// TwinCAT 3 PLC project slavePLC
// ProgramVersion: 3.1.4026.20
// libraries:
//   Tc2_Standard, * (Beckhoff Automation GmbH)
//   Tc2_System, * (Beckhoff Automation GmbH)
//   Tc3_Module, * (Beckhoff Automation GmbH)
//   VisuSymbols,3.5.10.0,System
// project tree:
//   / GlobalTextList.TcGTLO, PlcTask.TcTTO, Visualization Manager.TcVMO (not stored)
//   GVLs/ GVLSlave.TcGVL, ImagePoolCar.TcIPO (not stored)
//   POUs/ CarContorl.TcPOU, LampDelay.TcPOU, LampSlave.TcPOU, LongHandshake.TcPOU, MAIN.TcPOU, RunSlave.TcPOU, ShortHandshake.TcPOU, SlaveHandeshake.TcPOU
//   VISUs/ VisualizationSlave.TcVIS
// (motion and I/O tree: see PLC project studentplc)
// real-time tasks:
//   TASK PlcTask: cycle T#10ms, priority 20, ADS port 350
//   TASK PlcTask1: cycle T#10ms, priority 21, ADS port 351
// variable links:
//   StudentPLC/StudentPLC Instance <-> slavePLC/slavePLC Instance
//     PlcTask Inputs/GVLStudent.ixStrobOne <-> PlcTask Outputs/GVLSlave.oxStrobOne
//     PlcTask Inputs/GVLStudent.ixStrobTwo <-> PlcTask Outputs/GVLSlave.oxStrobTwo
//     PlcTask Outputs/GVLStudent.IXButtonLong <-> PlcTask Inputs/GVLSlave.ixLong
//     PlcTask Outputs/GVLStudent.IXButtonShort <-> PlcTask Inputs/GVLSlave.ixShort
//     PlcTask Outputs/GVLStudent.oxStrobOne <-> PlcTask Inputs/GVLSlave.ixStrobOne
//     PlcTask Outputs/GVLStudent.oxStrobTwo <-> PlcTask Inputs/GVLSlave.ixStrobTwo

CONFIGURATION slavePLC
    RESOURCE PLC ON TwinCAT3
        TASK PlcTask(INTERVAL := T#10ms, PRIORITY := 21);
        PROGRAM MAIN WITH PlcTask : MAIN;
    END_RESOURCE
END_CONFIGURATION

// ---- GVLs/GVLSlave.TcGVL
{attribute 'qualified_only'}
VAR_GLOBAL
	
	// Lamp varibol
	OXLampOXOne :BOOL;
	OXLampIXOneGreen :BOOL;
	OXLampOXTwo :BOOL;
	OXLampIXTwoGreen :BOOL;
	
	//strob out
	oxStrobOne AT %Q* : BOOL ;
	oxStrobTwo AT %Q* : BOOL ;
 	//strob in
	ixStrobOne AT %I* : BOOL ;
	ixStrobTwo AT %I* : BOOL ;
	
	// Long or Short
	ixLong AT %I* : BOOL;
	ixShort AT%I* :BOOL;
	
	// car move
	OIntRedCar: INT;
	OintCopCar: INT;
END_VAR

// ---- POUs/MAIN.TcPOU
PROGRAM MAIN
VAR
END_VAR

RunSlave();

END_PROGRAM

// ---- POUs/RunSlave.TcPOU
PROGRAM RunSlave
VAR
	LampSlave_0: LampSlave;
	SlaveHandeshake_0: SlaveHandeshake;
	ixStrobOne :BOOL;
	ixStrobTwo :BOOL;
	startCar: BOOL;
	carEnd: BOOL;
	CarContorl_0: CarContorl;
END_VAR

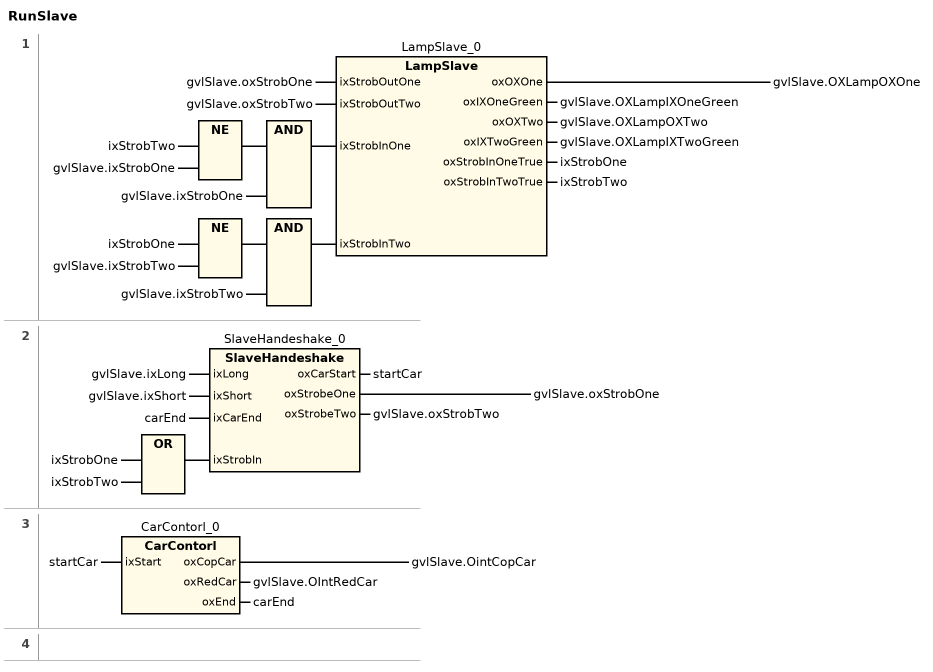
// NETWORK 1
LampSlave_0(
    ixStrobOutOne := gvlSlave.oxStrobOne,
    ixStrobOutTwo := gvlSlave.oxStrobTwo,
    ixStrobInOne := ixStrobTwo <> gvlSlave.ixStrobOne AND gvlSlave.ixStrobOne,
    ixStrobInTwo := ixStrobOne <> gvlSlave.ixStrobTwo AND gvlSlave.ixStrobTwo,
    oxIXOneGreen => gvlSlave.OXLampIXOneGreen,
    oxOXTwo => gvlSlave.OXLampOXTwo,
    oxIXTwoGreen => gvlSlave.OXLampIXTwoGreen,
    oxStrobInOneTrue => ixStrobOne,
    oxStrobInTwoTrue => ixStrobTwo); // LampSlave
gvlSlave.OXLampOXOne := LampSlave_0.oxOXOne;

// NETWORK 2
SlaveHandeshake_0(
    ixLong := gvlSlave.ixLong,
    ixShort := gvlSlave.ixShort,
    ixCarEnd := carEnd,
    ixStrobIn := ixStrobOne OR ixStrobTwo,
    oxCarStart => startCar,
    oxStrobeTwo => gvlSlave.oxStrobTwo); // SlaveHandeshake
gvlSlave.oxStrobOne := SlaveHandeshake_0.oxStrobeOne;

// NETWORK 3
CarContorl_0(ixStart := startCar, oxRedCar => gvlSlave.OIntRedCar, oxEnd => carEnd); // CarContorl
gvlSlave.OintCopCar := CarContorl_0.oxCopCar;

// NETWORK 4

END_PROGRAM

// ---- POUs/LampSlave.TcPOU
FUNCTION_BLOCK LampSlave
VAR_INPUT
	ixStrobOutOne :BOOL; // Direct control for group One main lamp (OX1)
	ixStrobOutTwo :BOOL; // Direct control for group Two main lamp (OX2)
	
	ixStrobInOne: BOOL; // Start signal for LampDelay sequence (group One)
	ixStrobInTwo: BOOL; // Start signal for LampDelay sequence (group Two)

END_VAR
VAR_OUTPUT
	  // Group One: main lamp + 3 indicator lamps (R, B, G)
	oxOXOne :BOOL; // Main lamp (direct)
	
	oxIXOneGreen :BOOL; // Indicator Green (from LampDelay)
	
	oxOXTwo :BOOL; // Main lamp (direct)
	
	oxIXTwoGreen :BOOL; // Indicator Green (from LampDelay)
	
	oxStrobInOneTrue: BOOL; // TRUE when all three indicators (group One) are ON
	oxStrobInTwoTrue: BOOL;// TRUE when all three indicators (group Two) are ON
	
END_VAR
	
VAR
	
	LampIXOne : LampDelay; // Instance for group One sequence
	LampIXTwo : LampDelay; // Instance for group Two sequence
	
END_VAR

// ------------------------------
// Direct main-lamp control
// ------------------------------

IF ixStrobOutOne THEN
	oxOXOne := TRUE;
ELSE
	oxOXOne := FALSE;
END_IF

IF ixStrobOutTwo THEN
	oxOXTwo := TRUE;
ELSE
	oxOXTwo := FALSE;
END_IF



// ------------------------------
// Group One: delayed indicator sequence
// ------------------------------
LampIXOne(ixStart := ixStrobInOne);

// Map LampDelay outputs to group One indicators
oxIXOneGreen     := LampIXOne.oxLampThree; // Green
oxStrobInOneTrue := LampIXOne.oxAllLightsOn; // All indicators ON


// ------------------------------
// Group Two: delayed indicator sequence
// ------------------------------
LampIXTwo(ixStart := ixStrobInTwo);

// Map LampDelay outputs to group Two indicators
oxIXTwoGreen     := LampIXTwo.oxLampThree; // Green
oxStrobInTwoTrue := LampIXTwo.oxAllLightsOn; // All indicators ON

END_FUNCTION_BLOCK

// ---- POUs/LampDelay.TcPOU
FUNCTION_BLOCK LampDelay
VAR_INPUT
    ixStart : BOOL;      // Start command: TRUE = run "power-up" sequence; FALSE = run "power-down" sequence
END_VAR
VAR_OUTPUT
    oxLampThree    : BOOL; // Output: Lamp 3 on/off
    oxAllLightsOn  : BOOL; // TRUE when all three lamps are on
END_VAR
VAR
    t      : TON;             // TON timer instance (non-retentive on IN falling edge)
    step   : INT := 0;        // State machine step
    delay  : TIME := T#2S;    // Delay duration used between steps
    tStart : BOOL;            // Timer IN signal (acts like a "strobe" to start the TON)
    tEnd   : BOOL;            // TRUE when timer has elapsed (t.Q)
END_VAR


//_______________________________________________________________________________________________
// LampDelay is a step-sequenced (state machine) controller that turns on three lamps
// one BY one with a fixed delay between each stage when ixStart is TRUE. 
// When ixStart goes FALSE, it turns the lamps off again in reverse order, also with delays. 
// A TON timer (t) provides the per-step delay. oxAllLightsOn is TRUE once all three lamps are on.
//_______________________________________________________________________________________________


// ------------------------------
// State machine for sequenced on/off with delays
// ------------------------------
CASE step OF

    0: // Idle/reset: all lamps off, wait for start
        oxLampThree    := FALSE;
        oxAllLightsOn  := FALSE;
        IF ixStart THEN
            // Start power-up sequence: immediately turn on Lamp 1 and start delay
            tStart    := TRUE;                  // Start the TON for the next step delay
			t(IN := tStart, PT := delay);
            step      := 20;
        END_IF


    20: // After Lamp 2 is on, wait delay, then turn on Lamp 3
        IF tEnd THEN
            tStart := FALSE;                   // Reset TON input before next start
            t(IN := tStart, PT := delay);
            oxLampThree := TRUE;
            step := 30;
        END_IF

    30: // All three lamps are on; assert "all on" and wait for stop command
        oxAllLightsOn := TRUE;
        IF NOT ixStart THEN
            // Begin power-down sequence after stop command
            tStart := TRUE;                    // Start delay before turning lamps off
            t(IN := tStart, PT := delay);
            step := 60;
        END_IF


    60: // Wait delay, then turn off Lamp 1 and return to idle
        IF tEnd THEN
            oxLampThree := FALSE;
			tStart := FALSE;
			t(IN := tStart,  PT := delay);
            step := 0;                         // Back to idle
        END_IF

END_CASE

// ------------------------------
// Timer execution (must be called each cycle)
// ------------------------------
t(IN := tStart, PT := delay);  // Evaluate TON with current IN/PT
tEnd := t.Q;                   // Timer done flag for step logic

END_FUNCTION_BLOCK

// ---- POUs/SlaveHandeshake.TcPOU
FUNCTION_BLOCK SlaveHandeshake
VAR_INPUT
	ixLong :BOOL;
	ixShort :BOOL;
	ixCarEnd: BOOL;
	ixStrobIn :BOOL; 
END_VAR
VAR_OUTPUT
	oxCarStart: BOOL;
	oxStrobeOne : BOOL;
    oxStrobeTwo : BOOL;
END_VAR
VAR
	
	long : LongHandshake;
	short : ShortHandshake;  
	oxStrobeOneShort : BOOL;
	oxStrobeOneLong : BOOL;
	oxCarStartLong: BOOL;
	oxCarStartShort: BOOL;
	step : INT := 0;
	waitLong : BOOL;
	waitShort: BOOL;
END_VAR

// ------------------------------
// State selector: choose which handshake to run
// ------------------------------
CASE step OF

    0: // IDLE: wait for a mode selection
        // NOTE: If both ixLong and ixShort are TRUE, long wins here.
        IF ixLong THEN
            step := 10;
        ELSIF ixShort THEN
            step := 20;
        END_IF

    10: // RUN LONG HANDSHAKE
        long(ixStart := ixCarEnd, ixStrobIn := ixStrobIn);

        // Map long handshake outputs to locals
        oxStrobeOneLong := long.oxStrobeOne;
        oxStrobeTwo     := long.oxStrobeTwo;  // direct passthrough (long only)
        oxCarStartLong  := long.oxStart;
        waitLong        := long.oxwait;

        // When long handshake reports idle, return to IDLE
        IF waitLong THEN
            step := 0;
        END_IF

    20: // RUN SHORT HANDSHAKE
        short(ixStart := ixCarEnd, ixStrobIn := ixStrobIn);

        // Map short handshake outputs to locals
        oxStrobeOneShort := short.oxStrobe;
        oxCarStartShort  := short.oxStart;
        waitShort        := short.oxwait;     // FIX: lowercase 'short'

        // When short handshake reports idle, return to IDLE
        IF waitShort THEN
            step := 0;
        END_IF

END_CASE


// ------------------------------
// Common output mapping
// ------------------------------

// Car start/ack goes TRUE if either handshake asserts it
IF oxCarStartShort OR oxCarStartLong THEN 
	oxCarStart := TRUE; 
ELSE 
	oxCarStart := FALSE; 
END_IF

// Primary strobe is TRUE if either handshake asserts it
IF oxStrobeOneShort OR oxStrobeOneLong THEN
	oxStrobeOne := TRUE; 
ELSE 
	oxStrobeOne := FALSE; 
END_IF

END_FUNCTION_BLOCK

// ---- POUs/LongHandshake.TcPOU
FUNCTION_BLOCK LongHandshake
VAR_INPUT
    ixStart   : BOOL; // From Master: start command ("execute now")
    ixStrobIn : BOOL; // From Master: strobe/ack line used through the long handshake
END_VAR
VAR_OUTPUT
    oxStart     : BOOL; // To Master: Slave "start request" (go-high to request start)
    oxStrobeOne : BOOL; // To Master: first Slave strobe (ack for initial Master strobe)
    oxStrobeTwo : BOOL; // To Master: second Slave strobe (ack after start)
    oxwait      : BOOL; // TRUE when idle/waiting; FALSE during handshake
END_VAR
VAR
    step : INT := 0;     // State machine step
END_VAR

CASE step OF

    0:  // IDLE: reset strobes, signal wait, and watch for Master strobe
        oxStrobeOne := FALSE;
        oxStrobeTwo := FALSE;
        oxStart     := FALSE;   // Ensure start request is low in idle
        oxwait      := TRUE;

        IF ixStrobIn THEN
            // Master raised strobe → acknowledge with Slave strobe one
            oxStrobeOne := TRUE;
            oxwait      := FALSE;
            step        := 10;
        END_IF

    10: // HOLD STROBE ONE until Master drops its strobe
        oxStrobeOne := TRUE;

        IF NOT ixStrobIn THEN
            // Master dropped strobe → drop Slave strobe one and move on
            oxStrobeOne := FALSE;
            step        := 20;
        END_IF

    20: // REQUEST START: raise oxStart to ask Master to start
        oxStart := TRUE;        // Keep high until Master issues ixStart

        IF ixStart THEN
            // Start received → drop request and raise second strobe
            oxStart     := FALSE;
            oxStrobeTwo := TRUE;
            step        := 30;
        END_IF

    30: // HOLD STROBE TWO until Master acknowledges (raises its strobe)
        oxStrobeTwo := TRUE;

        IF ixStrobIn THEN
            // Master acknowledged → drop strobe two and wait for final low
            oxStrobeTwo := FALSE;
            step        := 40;
        END_IF

    40: // WAIT FOR MASTER TO RETURN LOW to complete the cycle
        oxStrobeTwo := FALSE;

        IF NOT ixStrobIn THEN
            // Handshake finished → back to idle
            step := 0;
        END_IF

END_CASE

END_FUNCTION_BLOCK

// ---- POUs/ShortHandshake.TcPOU
FUNCTION_BLOCK ShortHandshake
VAR_INPUT
    ixStart   : BOOL; // Input from Master: start command ("execute now")
    ixStrobIn : BOOL; // Input from Master: strobe/trigger to initiate the handshake
END_VAR

VAR_OUTPUT
    oxStart  : BOOL; // Output to Master: "acknowledge/ready" from Slave
    oxStrobe : BOOL; // Output to Master: Slave strobe/confirmation during handshake
    oxwait   : BOOL; // Output: TRUE when Slave is idle/waiting
END_VAR

VAR
    step : INT := 0; // State machine step
END_VAR


// ------------------------------
// Short handshake sequence (Slave side)
// Step 0: Idle, waiting for Master strobe (ixStrobIn = TRUE)
// Step 10: Acknowledge/ready (oxStart = TRUE) until Master issues start (ixStart = TRUE)
// Step 20: Slave strobe (oxStrobe = TRUE) until Master drops its strobe (ixStrobIn = FALSE)
// ------------------------------
CASE step OF

    0:  // IDLE: reset all signals, wait for Master strobe
        oxStrobe := FALSE;
        oxStart  := FALSE;
        oxwait   := TRUE;

        IF ixStrobIn THEN
            // Master raised strobe → acknowledge and go to READY
            oxStart := TRUE;
            oxwait  := FALSE;
            step    := 10;
        END_IF

    10: // READY: wait for Master start command
        oxStart := TRUE;   // Keep acknowledge high

        IF ixStart THEN
            // Master gave start → drop ack and raise Slave strobe
            oxStart  := FALSE;
            oxStrobe := TRUE;
            step     := 20;
        END_IF

    20: // SLAVE STROBE: hold until Master drops its strobe
        oxStrobe := TRUE;

        IF NOT ixStrobIn THEN
            // Master strobe dropped → finish cycle and return to idle
            oxStrobe := FALSE;
            step     := 0;
        END_IF

END_CASE

END_FUNCTION_BLOCK

// ---- POUs/CarContorl.TcPOU
FUNCTION_BLOCK CarContorl
VAR_INPUT
    ixStart : BOOL;         // Start signal: TRUE = run sequence, FALSE = reset
END_VAR
VAR_OUTPUT
    oxCopCar : INT;         // Position counter for Cop car (moves negative)
    oxRedCar : INT;         // Position counter for Red car (moves negative)
    oxEnd    : BOOL;        // TRUE when both cars reach their thresholds
END_VAR
VAR
    step   : INT := 0;      // Step in the state machine
    t      : TON;           // TON timer instance (1s delay)
    delay  : TIME := T#1S;  // Delay interval
    tStart : BOOL;          // TON input (used as strobe to retrigger timer)
    tEnd   : BOOL;          // TON output (TRUE when delay time has passed)
END_VAR

//_______________________________________________________________________________________________________________
// CarContorl is a simple state machine that simulates two “cars” moving when the start signal (ixStart) is TRUE.
// Every second, the Cop car counter decreases by 2 and the Red car counter decreases by 3.
// When both cars pass their thresholds (Cop ≤ −800 and Red ≤ −1000), the output oxEnd is set TRUE.
// If ixStart goes FALSE, everything resets to the initial state.
//______________________________________________________________________________________________________________

CASE step OF

    0:  // IDLE/RESET: clear outputs and wait for start
        oxEnd    := FALSE;
        oxCopCar := 0;
        oxRedCar := 0;

        IF ixStart THEN
            tStart := TRUE;                // Start the first delay
            t(IN := tStart, PT := delay);
            step := 1;
        END_IF

    1:  // UPDATE POSITION: decrement both cars each cycle
        oxCopCar := oxCopCar - 2;          // Cop car moves -2 per step
        oxRedCar := oxRedCar - 3;          // Red car moves -3 per step

        IF tEnd THEN                       // After 1 second → go to check
            step := 10;
        END_IF

    10: // CHECK GOALS: have both thresholds been reached?
        IF (oxCopCar <= -800) AND (oxRedCar <= -1000) THEN
            oxEnd := TRUE;                 // Both goals reached → finish
            step  := 20;
        ELSE
            // Not yet → retrigger TON for next cycle
            tStart := FALSE;               // Reset TON input
            t(IN := tStart, PT := delay);
            tStart := TRUE;                // Rising edge to retrigger TON
            t(IN := tStart, PT := delay);
            step := 1;                     // Continue updating
        END_IF

    20: // FINISHED: hold end signal until start goes low
        oxEnd := TRUE;

        IF NOT ixStart THEN                // Stop command → reset
            oxEnd := FALSE;
            step  := 0;
        END_IF

END_CASE

// ------------------------------
// Timer evaluation – must be called every cycle
// ------------------------------
t(IN := tStart, PT := delay);
tEnd := t.Q;

END_FUNCTION_BLOCK

// ---- GlobalTextList.TcGTLO
TEXTLIST GlobalTextList
  76 = "first strobe '\\n' downloaded"
  36 = 'first strobe downloaded'
  378 = 'IXOne'
  620 = 'IXTwo'
  958 = 'loading'
  923 = 'Looding'
  389 = 'Loodining'
  816 = 'OXOne'
  99 = 'OXTwo'
  160 = 'Slav PLC'
  965 = 'Slav Strob One '
  171 = 'Slav strob one send'
  590 = 'Slav strob Two send'
  605 = 'Slav strob two send'
  659 = 'Strob sent'
  46 = 'strobe downloaded'
  781 = 'Strobe downloaded'
  391 = 'strobe received'
  968 = 'Strobe received'
END_TEXTLIST

// ---- VISUs/VisualizationSlave.TcVIS
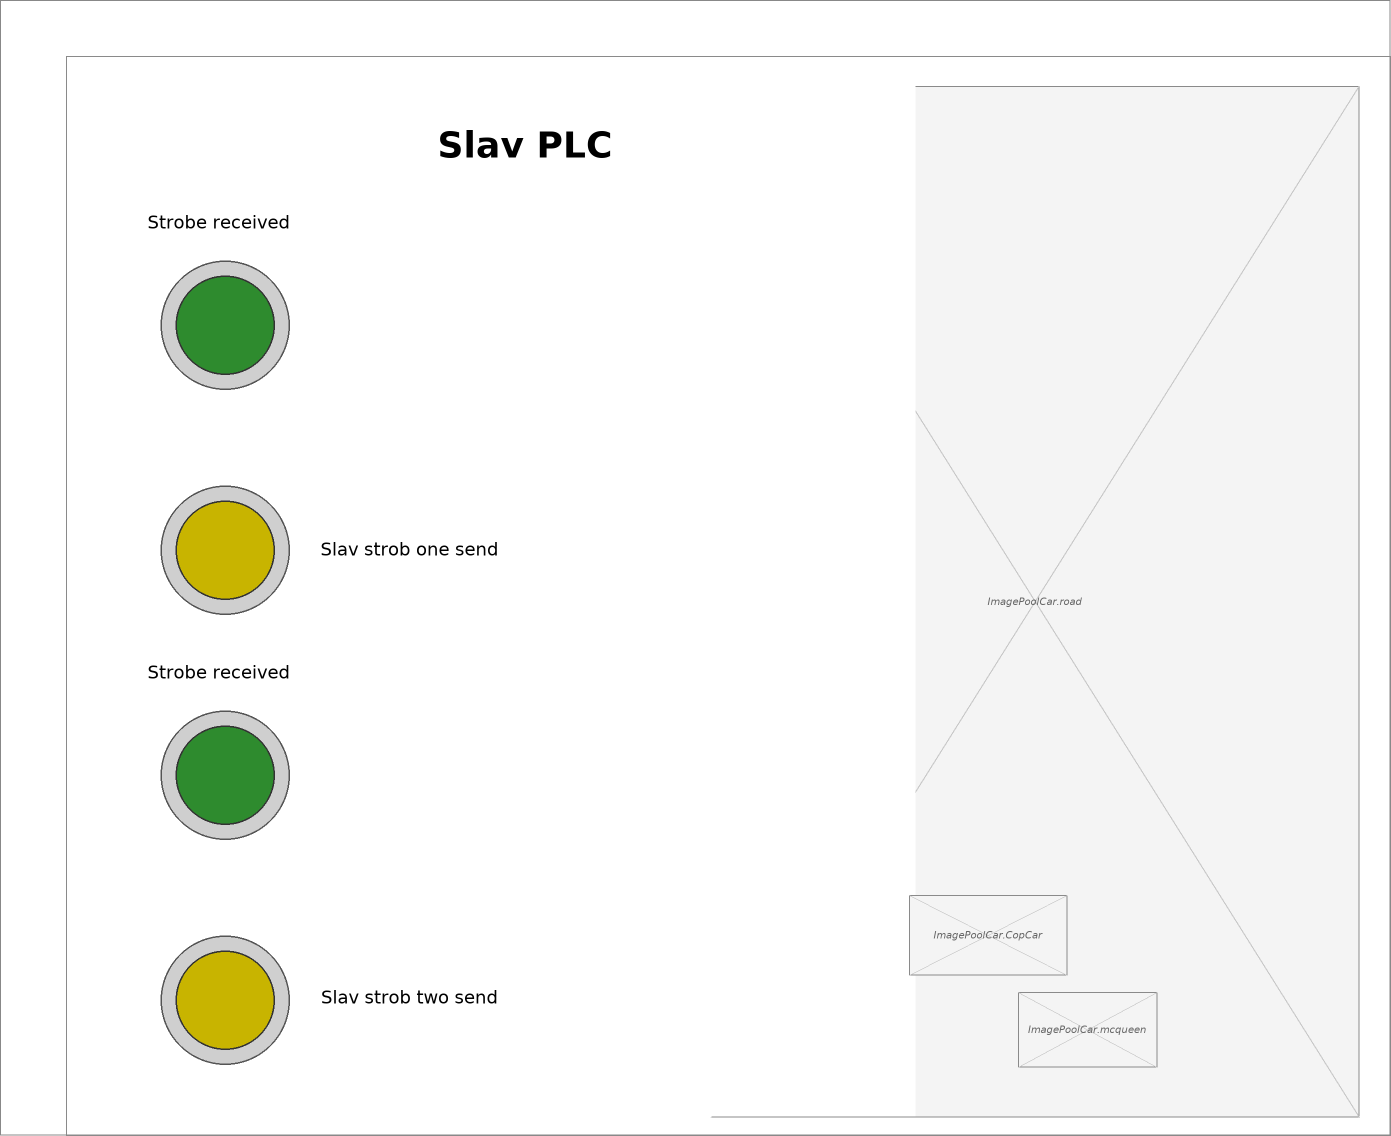
VISUALIZATION VisualizationSlave  // 1391x1136
    Frame (66,56 1325x1080)
    Image (711,86 648x1031), image: ImagePoolCar.road
    Rectangle (637,86 278x1030)
    Label (400,120 250x50), "Slav PLC"
    Lamp1 (150,250 150x150), variable: GVLSlave.OXLampIXOneGreen, style: Lamp-Lamp1-Green
    Label (100,200 238x45), "Strobe received"
    Label (300,527 219x45), "Slav strob one send"
    Lamp1 (150,475 150x150), variable: GVLSlave.OXLampOXOne, style: Lamp-Lamp1-Yellow
    Lamp1 (150,700 150x150), variable: GVLSlave.OXLampIXTwoGreen, style: Lamp-Lamp1-Green
    Lamp1 (150,925 150x150), variable: GVLSlave.OXLampOXTwo, style: Lamp-Lamp1-Yellow
    Image (1018,992 139x75), angle 90, image: ImagePoolCar.mcqueen
        p3528305787: GVLSlave.OIntRedCar
        p874137650: GVLSlave.OIntRedCar
    Image (909,895 158x80), angle 90, image: ImagePoolCar.CopCar
        p3528305787: GVLSlave.OintCopCar
        p874137650: GVLSlave.OintCopCar
    Label (300,975 219x45), "Slav strob two send"
    Label (100,650 238x45), "Strobe received"
    Label (450,650 150x30)
END_VISUALIZATION
